Fanuc KAREL source: KA00128.KL

PROGRAM KA00128
%NOLOCKGROUP
VAR
  SRC: ARRAY[2] OF BYTE
  DST: JOINTPOS
BEGIN
  SRC[1] = 2
  DST = SRC[1]
END KA00128
